(* IEC 61131-3 sources: kns-port-domestic/tools/port_metrics_tests/fixtures/adapted/src/POUs/FB_Pump, 3 files *)

(* ---- FB_Pump.decl.st ---- *)
// Насос: пример для метрик переноса
// PORT: [oop] EXTENDS не подтверждён в Astra.IDE (F23) — база вложена экземпляром
FUNCTION_BLOCK FB_Pump
VAR_INPUT
    xStart : BOOL;
    stCfg : ST_PumpCfg;
END_VAR
VAR_OUTPUT
    xRunning : BOOL;
END_VAR
VAR
    tonDelay : TON;
    fbBase : FB_Base; // PORT: [oop] композиция вместо наследования
END_VAR

(* ---- FB_Pump.impl.st ---- *)
// PORT: [oop] вызов базы через экземпляр вместо SUPER^
fbBase();
tonDelay(IN := xStart, PT := stCfg.tStartDelay);
xRunning := tonDelay.Q AND NOT fbBase.xFault; // PORT: доступ к полю базы через экземпляр (наследование)
IF xRunning THEN
    Start();
ELSE
    Stop();
END_IF

(* ---- Start.method.decl.st ---- *)
METHOD Start : BOOL
VAR_INPUT
END_VAR
